// TIA Portal V21 export
// export: Created 2026-11-10T07:35:18.4160664Z, ExportSetting WithDefaults, DisplayName Totally Integrated Automation Portal, DisplayVersion V21 Update 3, DisplayName STEP 7 Professional, DisplayVersion V21 Update 3, DisplayName STEP 7 Safety, DisplayVersion V21, DisplayName Tech WebApplication, DisplayVersion V21, DisplayName WinCC Basic/Comfort/Advanced, DisplayVersion V21 Update 3, DisplayName WinCC Unified, DisplayVersion V21 Update 3
FUNCTION_BLOCK "FB_Lad_ex133"   // FB52, LAD
{ S7_Optimized_Access := 'TRUE' }
VERSION : 0.1
// stored: AutoNumber true, IsIECCheckEnabled false, IsRetainMemResEnabled false, MemoryReserve 100, SetENOAutomatically false, UDAEnableTagReadback false
   VAR_INPUT
      v_mode : UInt;
      v_laddr : HW_ANY;
      v_ret_val : Int;
   END_VAR
   VAR_OUTPUT
      v_cnt_diag : UInt;
   END_VAR
   VAR_IN_OUT
      v_diag : Variant;
      v_detail : Variant;
   END_VAR
BEGIN

REGION Network 1: GET_DIAG - Read diagnostic information
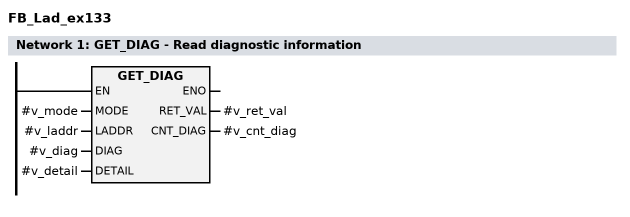
   RUNG wire#powerrail
      GET_DIAG(MODE := #v_mode, LADDR := #v_laddr, RET_VAL => #v_ret_val, CNT_DIAG => #v_cnt_diag, DIAG := #v_diag, DETAIL := #v_detail)
   END_RUNG
   // the same network as SCL:
   #v_ret_val := GET_DIAG(MODE := #v_mode,
                          LADDR := #v_laddr,
                          DIAG := #v_diag,
                          DETAIL := #v_detail,
                          CNT_DIAG => #v_cnt_diag);
END_REGION
END_FUNCTION_BLOCK
